(* IEC 61131-3 sources: openplc-editor-canopen/e2e/fixtures/cpp-compile-error/pous/programs, 1 file *)

(* ---- main.st ---- *)
PROGRAM main
  VAR
    counter : DINT;
    block : cpp_fb;
  END_VAR

counter := counter + 1;
block(in_val := counter);

END_PROGRAM
